(* IEC 61131-3 sources: plcassist-cli/packages/volt-lsp-iec/test-corpus/bakon-nano/Device/Plc Logic/Application/Library Manager/CmpDynamicText, 22 files *)

(* ---- DYNAMICTEXTCHANGELANGUAGE.fun ---- *)
FUNCTION DYNAMICTEXTCHANGELANGUAGE : BOOL
VAR_INPUT
	STLANGUAGE : STRING;
END_VAR
END_FUNCTION

(* ---- DYNAMICTEXTGETCURRENTLANGUAGE.fun ---- *)
FUNCTION DYNAMICTEXTGETCURRENTLANGUAGE : STRING
END_FUNCTION

(* ---- DYNAMICTEXTGETDEFAULTTEXT.fun ---- *)
FUNCTION DYNAMICTEXTGETDEFAULTTEXT : POINTER TO STRING
VAR_INPUT
	PSTTEXTLIST : POINTER TO STRING;
	PSTTEXTINDEX : POINTER TO STRING;
END_VAR
END_FUNCTION

(* ---- DYNAMICTEXTGETDEFAULTTEXTW.fun ---- *)
FUNCTION DYNAMICTEXTGETDEFAULTTEXTW : POINTER TO STRING
VAR_INPUT
	PSTTEXTLIST : POINTER TO STRING;
	PSTTEXTINDEX : POINTER TO STRING;
END_VAR
END_FUNCTION

(* ---- DYNAMICTEXTGETLANGUAGETEXT.fun ---- *)
FUNCTION DYNAMICTEXTGETLANGUAGETEXT : POINTER TO STRING
VAR_IN_OUT
	STLANGUAGE : STRING;
	STTEXTLIST : STRING;
	STTEXTINDEX : STRING;
END_VAR
END_FUNCTION

(* ---- DYNAMICTEXTGETLANGUAGETEXTW.fun ---- *)
FUNCTION DYNAMICTEXTGETLANGUAGETEXTW : POINTER TO WSTRING
VAR_IN_OUT
	STLANGUAGE : STRING;
	STTEXTLIST : STRING;
	STTEXTINDEX : STRING;
END_VAR
END_FUNCTION

(* ---- DYNAMICTEXTGETTEXT.fun ---- *)
FUNCTION DYNAMICTEXTGETTEXT : POINTER TO STRING
VAR_INPUT
	PSTTEXTLIST : POINTER TO STRING;
	PSTTEXTINDEX : POINTER TO STRING;
END_VAR
END_FUNCTION

(* ---- DYNAMICTEXTGETTEXTW.fun ---- *)
FUNCTION DYNAMICTEXTGETTEXTW : POINTER TO STRING
VAR_INPUT
	PSTTEXTLIST : POINTER TO STRING;
	PSTTEXTINDEX : POINTER TO STRING;
END_VAR
END_FUNCTION

(* ---- DYNAMICTEXTITERATEINDICES.fun ---- *)
FUNCTION DYNAMICTEXTITERATEINDICES : RTS_IEC_RESULT
VAR_INPUT
	PSTTEXTLIST : POINTER TO STRING;
	PFITERATIONCALLBACK : POINTER TO BYTE;
	ITERATIONDATA : __UXINT;
END_VAR
END_FUNCTION

(* ---- DYNAMICTEXTITERATELANGUAGES.fun ---- *)
FUNCTION DYNAMICTEXTITERATELANGUAGES : RTS_IEC_RESULT
VAR_INPUT
	PFITERATIONCALLBACK : POINTER TO BYTE;
	ITERATIONDATA : __UXINT;
END_VAR
END_FUNCTION

(* ---- DYNAMICTEXTLOADDEFAULTTEXTS.fun ---- *)
FUNCTION DYNAMICTEXTLOADDEFAULTTEXTS : RTS_IEC_RESULT
END_FUNCTION

(* ---- DYNAMICTEXTLOADLANGUAGE.fun ---- *)
FUNCTION DYNAMICTEXTLOADLANGUAGE : RTS_IEC_RESULT
VAR_INPUT
	STLANGUAGE : STRING;
END_VAR
END_FUNCTION

(* ---- DYNAMICTEXTREGISTERFILE.fun ---- *)
FUNCTION DYNAMICTEXTREGISTERFILE : RTS_IEC_RESULT
VAR_INPUT
	SZFILE : REFERENCE TO STRING;
END_VAR
END_FUNCTION

(* ---- DYNAMICTEXTREGISTERPATH.fun ---- *)
FUNCTION DYNAMICTEXTREGISTERPATH : RTS_IEC_RESULT
VAR_INPUT
	SZPATH : REFERENCE TO STRING;
END_VAR
END_FUNCTION

(* ---- DYNAMICTEXTRELEASELANGUAGES.fun ---- *)
FUNCTION DYNAMICTEXTRELEASELANGUAGES : RTS_IEC_RESULT
VAR_INPUT
	XFORCERELEASE : BOOL;
END_VAR
END_FUNCTION

(* ---- DYNAMICTEXTRELEASELOCK.fun ---- *)
FUNCTION DYNAMICTEXTRELEASELOCK : BOOL
END_FUNCTION

(* ---- DYNAMICTEXTRELOADTEXTS.fun ---- *)
FUNCTION DYNAMICTEXTRELOADTEXTS : RTS_IEC_RESULT
END_FUNCTION

(* ---- DYNAMICTEXTSETLOCK.fun ---- *)
FUNCTION DYNAMICTEXTSETLOCK : BOOL
END_FUNCTION

(* ---- DYNAMICTEXTTESTANDSETLOCK.fun ---- *)
FUNCTION DYNAMICTEXTTESTANDSETLOCK : BOOL
END_FUNCTION

(* ---- DYNAMICTEXTUNLOADLANGUAGE.fun ---- *)
FUNCTION DYNAMICTEXTUNLOADLANGUAGE : RTS_IEC_RESULT
VAR_INPUT
	STLANGUAGE : STRING;
END_VAR
END_FUNCTION

(* ---- DYNAMICTEXTUNREFERENCELANGUAGE.fun ---- *)
FUNCTION DYNAMICTEXTUNREFERENCELANGUAGE : RTS_IEC_RESULT
VAR_INPUT
	STLANGUAGE : STRING;
END_VAR
END_FUNCTION

(* ---- DYNAMICTEXTUNREGISTERFILE.fun ---- *)
FUNCTION DYNAMICTEXTUNREGISTERFILE : RTS_IEC_RESULT
VAR_INPUT
	SZFILE : REFERENCE TO STRING;
END_VAR
END_FUNCTION
